(* IEC 61131-3 sources: nautilus/cmd/naut/testdata/agents-md, 1 file *)

(* ---- scaling.st ---- *)
PROGRAM Scaling
(* Level in percent from the raw 4-20 mA signal, held to 0-100. *)
VAR
  pct : REAL;
END_VAR
pct := (LT101_Raw - 4.0) / 16.0 * 100.0;
IF pct < 0.0 THEN
  pct := 0.0;
END_IF;
IF pct > 100.0 THEN
  pct := 100.0;
END_IF;
LT101_Pct := pct;
END_PROGRAM
